(* IEC 61131-3 sources: Test-Git_ESME26/TestProgettoESME_26.fbsproj/TemplateFullProgrammingFramework_Migration.device.xml.v3^/Plc Logic.plclogic.xml.v3^/Application.application.xml.v3^/TemplateFullProgrammingFramework/Examples/ExampleModulesExtItf/SR_CharlyModuleExtItf.prg.st^, 1 file *)

(* ---- RegisterLoggerPoint.meth.st ---- *)
METHOD RegisterLoggerPoint
VAR_INPUT
	i_ifParent	: APL.IF_LoggerPoint;
	i_sName		: STRING[80];
END_VAR
VAR_OUTPUT
	q_etDiag	: GD.ET_Diag := GD.ET_Diag.Ok;
	q_etDiagExt	: ET_DiagExt := ET_DiagExt.Ok;
END_VAR

SR_CharlyModule.RegisterLoggerPoint(	i_ifParent	:= i_ifParent,
										i_sName		:= i_sName,
										q_etDiag	=> q_etDiag,
										q_etDiagExt	=> q_etDiagExt);
